// TwinCAT 3 PLC project Plc
// libraries:
//   Tc2_Standard, * (Beckhoff Automation GmbH)
// project tree:
//   POUs/ MAIN.TcPOU, FB_Fill.TcPOU, FB_Valve.TcPOU
//   DUTs/ ST_Recipe.TcDUT
//   GVLs/ GVL_Machine.TcGVL

// ---- DUTs/ST_Recipe.TcDUT
TYPE ST_Recipe :
STRUCT
	rTargetKg   : LREAL;
	rBulkCutoff : LREAL := 0.9;
	sName       : STRING(40);
END_STRUCT
END_TYPE

// ---- GVLs/GVL_Machine.TcGVL
{attribute 'qualified_only'}
VAR_GLOBAL
	nDrumsFilled : UDINT;
	bEStop AT %I* : BOOL;
END_VAR
VAR_GLOBAL CONSTANT
	MAX_MODULES : INT := 16;	// sizing constant: the runtime exports it without a READONLY flag
END_VAR

// ---- POUs/MAIN.TcPOU
PROGRAM MAIN
VAR
	fbFill      : FB_Fill;        // main filling sequence
	stRecipe    : ST_Recipe;
	nCycle      : UDINT;
	bStart AT %I* : BOOL;
END_VAR

nCycle := nCycle + 1;
fbFill(bEnable := bStart, stRecipe := stRecipe);
IF fbFill.bDone THEN
	GVL_Machine.nDrumsFilled := GVL_Machine.nDrumsFilled + 1;
END_IF

END_PROGRAM

// ---- POUs/FB_Fill.TcPOU
FUNCTION_BLOCK FB_Fill EXTENDS FB_Base
VAR_INPUT
	bEnable   : BOOL;
	stRecipe  : ST_Recipe;
END_VAR
VAR_OUTPUT
	bDone     : BOOL;
	bError    : BOOL;
END_VAR
VAR
	fbValve   : FB_Valve;         (* bulk valve *)
	fbFine    : FB_Valve;         (* fine valve *)
	eState    : E_FillState;
	tSettle   : TIME := T#500MS;
	arrWeights : ARRAY[0..9] OF LREAL;
END_VAR

CASE eState OF
	E_FillState.Idle:
		IF bEnable THEN eState := E_FillState.Bulk; END_IF
	E_FillState.Bulk:
		fbValve.Open();
END_CASE

METHOD Start : BOOL
VAR_INPUT
	rTarget : LREAL;
END_VAR
eState := E_FillState.Bulk;
Start := TRUE;
END_METHOD

END_FUNCTION_BLOCK

// ---- POUs/FB_Valve.TcPOU
FUNCTION_BLOCK FB_Valve
VAR_OUTPUT
	bOpen AT %Q* : BOOL;   // solenoid
END_VAR
VAR
	tOpened : TIME;
END_VAR

;

METHOD Open
bOpen := TRUE;
END_METHOD

PROPERTY IsOpen : BOOL
GET
IsOpen := bOpen;
END_GET
END_PROPERTY

END_FUNCTION_BLOCK
